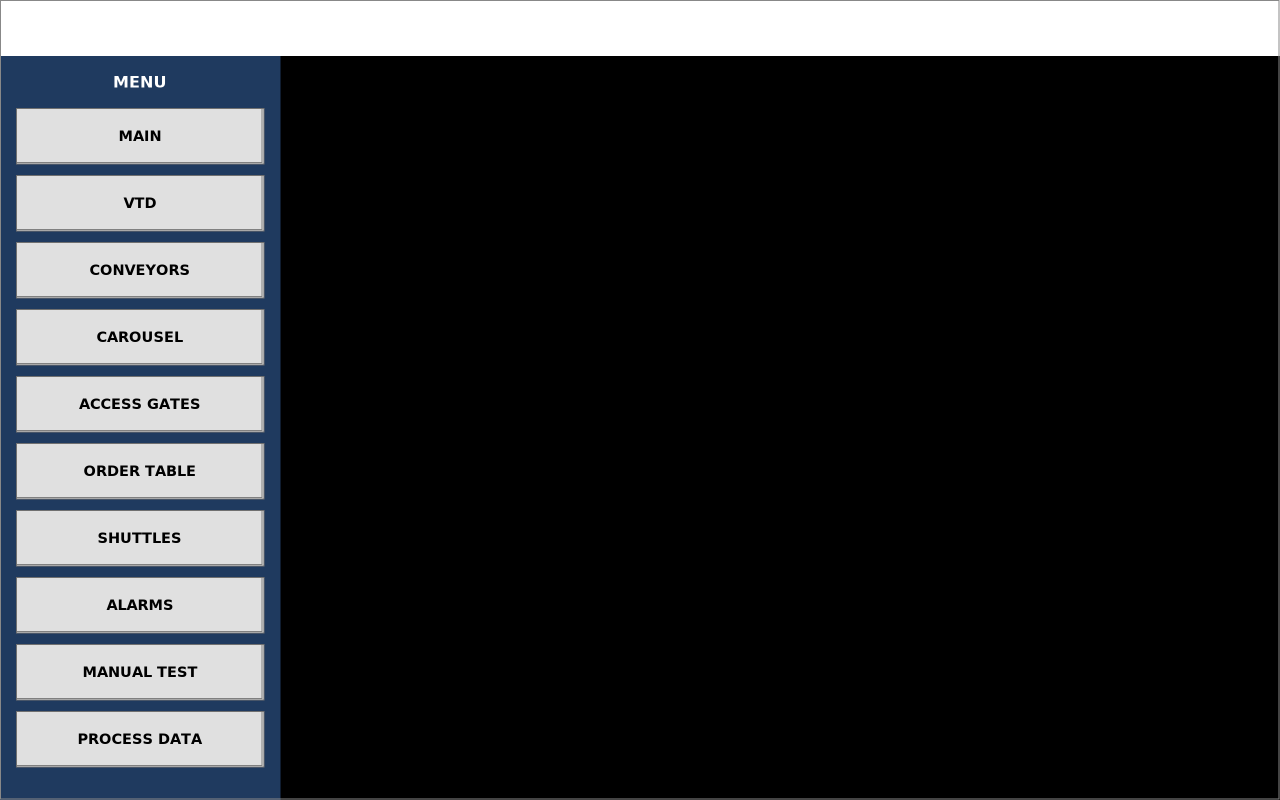
VISUALIZATION Dialog  // 1280x800
    Rectangle (0,0 1280x56)
        OnMouseClick: CloseDialog Dialog=Current Dialog, Result=OK, NumpadKeypadSet=True
    Rectangle (280,56 1000x744)
        OnMouseClick: CloseDialog Dialog=Current Dialog, Result=OK, NumpadKeypadSet=True
    Rectangle (0,56 280x744)
    Rectangle (12,64 256x36), "MENU"
    Button (16,108 248x56), "MAIN"
        OnMouseClick: CloseDialog Dialog=Current Dialog, Result=OK, NumpadKeypadSet=True
        OnMouseDown: change screen: Main
    Button (16,175 248x56), "VTD"
        OnMouseClick: CloseDialog Dialog=Current Dialog, Result=OK, NumpadKeypadSet=True
        OnMouseDown: change screen: VTD
    Button (16,242 248x56), "CONVEYORS"
        OnMouseClick: CloseDialog Dialog=Current Dialog, Result=OK, NumpadKeypadSet=True
        OnMouseDown: change screen: CNV
    Button (16,309 248x56), "CAROUSEL"
        OnMouseClick: CloseDialog Dialog=Current Dialog, Result=OK, NumpadKeypadSet=True
        OnMouseDown: change screen: Carrousel
    Button (16,376 248x56), "ACCESS GATES"
        OnMouseClick: CloseDialog Dialog=Current Dialog, Result=OK, NumpadKeypadSet=True
        OnMouseDown: change screen: Access_Gates
    Button (16,443 248x56), "ORDER TABLE"
        OnMouseClick: CloseDialog Dialog=Current Dialog, Result=OK, NumpadKeypadSet=True
        OnMouseDown: change screen: Order_Table
    Button (16,510 248x56), "SHUTTLES"
        OnMouseClick: CloseDialog Dialog=Current Dialog, Result=OK, NumpadKeypadSet=True
        OnMouseDown: change screen: Shuttles
    Button (16,577 248x56), "ALARMS"
        OnMouseClick: CloseDialog Dialog=Current Dialog, Result=OK, NumpadKeypadSet=True
        OnMouseDown: change screen: Alarms
    Button (16,644 248x56), "MANUAL TEST"
        OnMouseClick: CloseDialog Dialog=Current Dialog, Result=OK, NumpadKeypadSet=True
        OnMouseDown: change screen: VTDManualTest
    Button (16,711 248x56), "PROCESS DATA"
        OnMouseClick: CloseDialog Dialog=Current Dialog, Result=OK, NumpadKeypadSet=True
        OnMouseDown: change screen: Visualization
END_VISUALIZATION

(* stored: Version 1.1.0.1
   Visu Dialog: Id {8067e270-ca00-4168-8692-f5659e66b526} *)
